DATA_BLOCK "FRK_Profiles"
{ S7_Optimized_Access := 'TRUE' }
VERSION : 0.1
NON_RETAIN
VAR
    P001 {ExternalAccessible := 'False'; ExternalVisible := 'False'; ExternalWritable := 'False'} : "FRK_ProfileOwned_PressDemoUnit";
END_VAR
BEGIN
END_DATA_BLOCK
